(* IEC 61131-3 sources: XPGAnalyser/bac/Armoire_Gaz/ihm/fonctions, 2 files *)

(* ---- 0152-Moyenne_Pression.st ---- *)
(* Moyenne pondérée des pressions de deux armoires, en bar *)
VAR_INPUT
    A : REAL;
    B : REAL;
    Poids_A : REAL := 0.5;   (* 0.5 : la moyenne simple *)
END_VAR
VAR_TEMP
    Somme : REAL;
END_VAR

Somme := A * Poids_A + B * (1.0 - Poids_A);
Moyenne_Pression := Somme;

(* ---- 0153-Tracer_Evenement.st ---- *)
(* Une ligne au journal, et le compte des traces *)
VAR_INPUT
    Quoi : STRING;
    Niveau : INT := 1;
END_VAR

Compteur_Clics := Compteur_Clics + 1;
IF Niveau > 1 THEN
    IHM_JOURNAL('[ALERTE] {Quoi}');
ELSE
    IHM_JOURNAL('{Quoi}');
END_IF;
